(* IEC 61131-3 sources: Lasal-MCP/examples/SampleSource/LASALScreenAdvancedSolution/LASALScreenAdvancedSolution/LASALScreenAdvacnedSolution/Stations/Terminal/HMI/Class/MyScrollList, 1 file *)

(* ---- MyScrollList.st ---- *)
(*!
<Class
	Name               = "MyScrollList"
	Revision           = "0.0"
	RealtimeTask       = "false"
	CyclicTask         = "false"
	BackgroundTask     = "false"
	Sigmatek           = "false"
	OSInterface        = "false"
	HighPriority       = "false"
	Automatic          = "false"
	UpdateMode         = "Prescan"
	SharedCommandTable = "true"
	Objectsize         = "(540,240)">
	<Channels>
		<Client Name="_Grafix" Required="false" Internal="false"/>
		<Client Name="SigCLib" Required="false" Internal="false"/>
	</Channels>
	<Network Name="MyScrollList">
		<!-- List of Components in this network -->
		<Components>
			<Object
				Name       = "_base"
				Class      = "_ScrollArea2"
				Position   = "(218,120)"
				Visualized = "true"
				Remotely   = "true">
				<Channels>
					<Server Name="ActPos"/>
					<Server Name="Refresh"/>
					<Server Name="Server0"/>
					<Client Name="ExtendedScrollBar" Value="0"/>
					<Client Name="LineHighness"/>
					<Client Name="LineWidth"/>
					<Client Name="Lse"/>
					<Client Name="VerticalLevel"/>
				</Channels>
			</Object>
		</Components>
		<Comments>
		</Comments>
		<!-- List of Connections in this network -->
		<Connections>
			<Connection Source="this.Server0" Destination="_base.Server0" Vertices="(886,210),(714,210),"/>
			<Connection Source="this.Refresh" Destination="_base.Refresh" Vertices="(886,270),(714,270),"/>
			<Connection Source="this.ActPos" Destination="_base.ActPos" Vertices="(886,330),(714,330),"/>
			<Connection Source="_base.Lse" Destination="this.Lse" Vertices="(218,210),(38,210),"/>
			<Connection Source="_base.VerticalLevel" Destination="this.VerticalLevel" Vertices="(218,270),(38,270),"/>
			<Connection Source="_base.LineWidth" Destination="this.LineWidth" Vertices="(218,330),(38,330),"/>
		</Connections>
		<!-- Headerfiles -->
		<Options>
		</Options>
	</Network>
</Class>
*)
#pragma using _ScrollArea2

MyScrollList : CLASS
: _ScrollArea2
  //Servers:
  //Clients:
	_Grafix 	: CltChCmd__Grafix;
	SigCLib 	: CltChCmd_SigCLib;
  //Variables:
		pError 	: ^CHAR;
		intError 	: DINT;
  //Functions:

	FUNCTION VIRTUAL GLOBAL Init;
				//! <Function Comment="method is called every time when redraw of a single line is necessary.&#13;&#10;" Name="Line"/>
	FUNCTION __CDECL VIRTUAL GLOBAL Line
		VAR_INPUT
			ps 	: ^_SCROLL;			//! <Variable Comment="pointer to structure _SCROLL" Name="Line.ps"/>
			pr 	: ^_ROOM;			//! <Variable Comment="pointer to place where line should be drawn" Name="Line.pr"/>
			line 	: UINT;			//! <Variable Comment="16 bit linenumber " Name="Line.line"/>
			state 	: BOOL;			//! <Variable Comment="line is selected (true) or passive (false)" Name="Line.state"/>
		END_VAR;
  //Tables:
	FUNCTION @STD
		VAR_OUTPUT
			ret_code	: CONFSTATES;
		END_VAR;
	FUNCTION GLOBAL TAB @CT_;
END_CLASS;

#pragma usingLtd _Grafix
#pragma usingLtd SigCLib

FUNCTION VIRTUAL GLOBAL MyScrollList::Init
  // set Number of Lines
  if (_FirstScan = TRUE) then
    Scroll.position.no := 30;
  end_if;

END_FUNCTION

FUNCTION __CDECL VIRTUAL GLOBAL MyScrollList::Line
	VAR_INPUT
		ps 	: ^_SCROLL;
		pr 	: ^_ROOM;
		line 	: UINT;
		state 	: BOOL;
	END_VAR
  VAR
  	color : _COLOR;
    att : _ATTRIB;
    txt : array[0..29] of _ASCII;
  END_VAR

  // set color depending on state
  if (state = TRUE) then
    color := _Grafix.MakeColor(backcolor:= INVISIBLE,
                               frontcolor:= ps^.color_activ);
  else
    color := _Grafix.MakeColor(backcolor:= INVISIBLE,
                               frontcolor:= ps^.color_inactiv);

  end_if;

  // query on linenumber
  if (line < Scroll.position.no) then
    //set attributes
    att := T_LEFTBOUND or T_UPBOUND or T_COPY or T_PROP or T_SOLID;

    // column 1
    // --------------------------------------------------------------
    //copy string in array
    pError := SigCLib.StrCpy(dst0:= #txt[0],
                             src0:= "SIG-009-");

    if (pError <> #txt[0]) then
      intError := -1;
      return;
    end_if;

    //add linenumber to array
    DToA(p0:= #txt[8],
         x1:= line,
         x2:= 16#0800,
         x3:= sizeof(_ASCII));

    //draw string of first column
    _Grafix.OutTextXY(x0:= pr^.xy1.x + 10,
                      y0:= pr^.xy1.y,
                      textptr:= #txt[0],
                      attrib:= att,
                      color:= color,
                      chr_size:= sizeof(_ASCII));

    // column 2
    // --------------------------------------------------------------
    pError := SigCLib.StrCpy(dst0:= #txt[0],
                             src0:= "PR-X110-");

    if (pError <> #txt[0]) then
      intError := -2;
      return;
    end_if;

    txt[8] := 'A';
    txt[9] := 'A' + to_usint(line);
    txt[10] := 0;

    //draw string of second column
    _Grafix.OutTextXY(x0:= pr^.xy1.x + 200,
                      y0:= pr^.xy1.y,
                      textptr:= #txt[0],
                      attrib:= att,
                      color:= color,
                      chr_size:= sizeof(_ASCII));

    // column 3
    // --------------------------------------------------------------
    //draw string of third column
    _Grafix.OutTextXY(x0:= pr^.xy1.x + 400,
                      y0:= pr^.xy1.y,
                      textptr:= "Cat",
                      attrib:= att,
                      color:= color,
                      chr_size:= sizeof(_ASCII));

    //draw column seperator
    _Grafix.Line(x0:= pr^.xy1.x + 190,
                 y0:= pr^.xy1.y,
                 x1:= pr^.xy1.x + 190,
                 y1:= pr^.xy2.y,
                 attrib:= att,
                 color:= color);

    _Grafix.Line(x0:= pr^.xy1.x + 390,
                 y0:= pr^.xy1.y,
                 x1:= pr^.xy1.x + 390,
                 y1:= pr^.xy2.y,
                 attrib:= att,
                 color:= color);

  end_if;

END_FUNCTION
